PROGRAM MAIN
VAR
END_VAR

RunSlave();

END_PROGRAM

(* stored: Version 1.1.0.1, ProductVersion 3.1.4024.12
   POU MAIN: Id {a402e50a-06ad-425c-95ef-b54c55cf36ab}, SpecialFunc None *)
